(* IEC 61131-3 sources: plc-st-coding-agent/progress/evidence/f14_v11_public_20261113/jobs/codex_minimax-m27, 6 files *)

(* ---- public-easy-01.candidate_01.st ---- *)
(* ENGINEERING_CONTRACT
 * Filling Line State Machine - 6 states, sequential operation
 * PUB001: bottleSensor TRUE → Pump_Motor := TRUE (hold until cleaningConfirmButton)
 * PUB002: cleaningConfirmButton → Filling_Valve := TRUE (hold until fillingConfirmButton)
 * PUB003: fillingConfirmButton → Capping_Machine := TRUE (hold until cappingConfirmButton)
 * PUB004: cappingConfirmButton → Packing_Machine := TRUE (hold until packingConfirmButton)
 * PUB005: packingConfirmButton → Completion_Light := TRUE (hold until finishedButton)
 * PUB006: finishedButton → Completion_Light := FALSE; all outputs FALSE; reset to IDLE
 * State retention: outputs held until explicitly deactivated by state transition or reset
 * Reset priority: finishedButton (PUB006) clears all outputs and returns to IDLE
 *)

(* CONTRACT_RULES [] *)

FUNCTION_BLOCK FillingLineControl
VAR_INPUT
    bottleSensor          : BOOL;
    cleaningConfirmButton : BOOL;
    fillingConfirmButton  : BOOL;
    cappingConfirmButton  : BOOL;
    packingConfirmButton  : BOOL;
    finishedButton        : BOOL;
END_VAR
VAR_OUTPUT
    Pump_Motor      : BOOL;
    Filling_Valve   : BOOL;
    Capping_Machine : BOOL;
    Packing_Machine : BOOL;
    Completion_Light: BOOL;
END_VAR
VAR
    State : INT := 0;
END_VAR

// State machine: 0=IDLE, 1=CLEANING, 2=FILLING, 3=CAPPING, 4=PACKING, 5=COMPLETE
CASE State OF
    0: // IDLE - waiting for bottle
        Pump_Motor      := FALSE;
        Filling_Valve   := FALSE;
        Capping_Machine := FALSE;
        Packing_Machine := FALSE;
        Completion_Light:= FALSE;

        IF bottleSensor THEN
            State := 1;
        END_IF;

    1: // CLEANING
        Pump_Motor := TRUE;

        IF cleaningConfirmButton THEN
            Pump_Motor := FALSE;
            State := 2;
        END_IF;

    2: // FILLING
        Filling_Valve := TRUE;

        IF fillingConfirmButton THEN
            Filling_Valve := FALSE;
            State := 3;
        END_IF;

    3: // CAPPING
        Capping_Machine := TRUE;

        IF cappingConfirmButton THEN
            Capping_Machine := FALSE;
            State := 4;
        END_IF;

    4: // PACKING
        Packing_Machine := TRUE;

        IF packingConfirmButton THEN
            Packing_Machine := FALSE;
            State := 5;
        END_IF;

    5: // COMPLETE - bottle ready for pickup
        Completion_Light := TRUE;

        IF finishedButton THEN
            Completion_Light := FALSE;
            State := 0;
        END_IF;

END_CASE;

END_FUNCTION_BLOCK

(* ---- public-easy-01.raw_candidate_01.st ---- *)
(* ENGINEERING_CONTRACT
 * Filling Line State Machine - 6 states, sequential operation
 * PUB001: bottleSensor TRUE → Pump_Motor := TRUE (hold until cleaningConfirmButton)
 * PUB002: cleaningConfirmButton → Filling_Valve := TRUE (hold until fillingConfirmButton)
 * PUB003: fillingConfirmButton → Capping_Machine := TRUE (hold until cappingConfirmButton)
 * PUB004: cappingConfirmButton → Packing_Machine := TRUE (hold until packingConfirmButton)
 * PUB005: packingConfirmButton → Completion_Light := TRUE (hold until finishedButton)
 * PUB006: finishedButton → Completion_Light := FALSE; all outputs FALSE; reset to IDLE
 * State retention: outputs held until explicitly deactivated by state transition or reset
 * Reset priority: finishedButton (PUB006) clears all outputs and returns to IDLE
 *)

(* CONTRACT_RULES [] *)

FUNCTION_BLOCK FillingLineControl
VAR_INPUT
    bottleSensor          : BOOL;
    cleaningConfirmButton : BOOL;
    fillingConfirmButton  : BOOL;
    cappingConfirmButton  : BOOL;
    packingConfirmButton  : BOOL;
    finishedButton        : BOOL;
END_VAR
VAR_OUTPUT
    Pump_Motor      : BOOL;
    Filling_Valve   : BOOL;
    Capping_Machine : BOOL;
    Packing_Machine : BOOL;
    Completion_Light: BOOL;
END_VAR
VAR
    State : INT := 0;
END_VAR

// State machine: 0=IDLE, 1=CLEANING, 2=FILLING, 3=CAPPING, 4=PACKING, 5=COMPLETE
CASE State OF
    0: // IDLE - waiting for bottle
        Pump_Motor      := FALSE;
        Filling_Valve   := FALSE;
        Capping_Machine := FALSE;
        Packing_Machine := FALSE;
        Completion_Light:= FALSE;

        IF bottleSensor THEN
            State := 1;
        END_IF

    1: // CLEANING
        Pump_Motor := TRUE;

        IF cleaningConfirmButton THEN
            Pump_Motor := FALSE;
            State := 2;
        END_IF

    2: // FILLING
        Filling_Valve := TRUE;

        IF fillingConfirmButton THEN
            Filling_Valve := FALSE;
            State := 3;
        END_IF

    3: // CAPPING
        Capping_Machine := TRUE;

        IF cappingConfirmButton THEN
            Capping_Machine := FALSE;
            State := 4;
        END_IF

    4: // PACKING
        Packing_Machine := TRUE;

        IF packingConfirmButton THEN
            Packing_Machine := FALSE;
            State := 5;
        END_IF

    5: // COMPLETE - bottle ready for pickup
        Completion_Light := TRUE;

        IF finishedButton THEN
            Completion_Light := FALSE;
            State := 0;
        END_IF

END_CASE

END_FUNCTION_BLOCK

(* ---- public-easy-02.candidate_01.st ---- *)
(* ENGINEERING_CONTRACT
====================
PUB001: 76-318

State Retention:
- tmp_previous_value: RETAINED across scans (stores last cycle's DWORD value)
- All outputs: COMBINATIONAL (derived fresh each scan from current inputs + retained state)

Edge Detection Logic:
- Rising edge:  (current = 1) AND (previous = 0)  → risingBits = value & NOT previous
- Falling edge: (current = 0) AND (previous = 1)  → fallingBits = NOT value & previous
- Changed:      value <> previous

Counting:
- Count 1-bits in risingBits  → noOfRisingBits  (0-32)
- Count 1-bits in fallingBits → noOfFallingBits (0-32)

Priority:
- All outputs derived combinatorially in same scan
- No edge-only triggers or state machines

Units:
- risingBits/fallingBits: dimensionless bit patterns (DWORD)
- noOfRisingBits/noOfFallingBits: unsigned count (USINT, 0-32)
*)
FUNCTION_BLOCK FB_DualWordEdgeDetection
VAR
    tmp_previous_value : DWORD := 0;
END_VAR
VAR_OUTPUT
    hasChanged      : BOOL;
    hasRisingEdges  : BOOL;
    risingBits      : DWORD;
    noOfRisingBits  : USINT;
    hasFallingEdges : BOOL;
    fallingBits     : DWORD;
    noOfFallingBits : USINT;
END_VAR

risingBits  := value AND NOT tmp_previous_value;
fallingBits := NOT value AND tmp_previous_value;

hasChanged      := (value <> tmp_previous_value);
hasRisingEdges  := (risingBits <> 0);
hasFallingEdges := (fallingBits <> 0);

noOfRisingBits  := 0;
FOR i := 0 TO 31 DO
    IF SHR(risingBits, i) AND 1 = 1 THEN
        noOfRisingBits := noOfRisingBits + 1;
    END_IF;
END_FOR;

noOfFallingBits := 0;
FOR i := 0 TO 31 DO
    IF SHR(fallingBits, i) AND 1 = 1 THEN
        noOfFallingBits := noOfFallingBits + 1;
    END_IF;
END_FOR;

tmp_previous_value := value;
END_FUNCTION_BLOCK

(* ---- public-easy-02.candidate_02.st ---- *)
(* ENGINEERING_CONTRACT
====================
PUB001: 76-318

State Retention:
- tmp_previous_value: RETAINED across scans (stores last cycle's DWORD value)
- All outputs: COMBINATIONAL (derived fresh each scan from current inputs + retained state)

Edge Detection Logic:
- Rising edge:  (current = 1) AND (previous = 0)  → risingBits = value & NOT previous
- Falling edge: (current = 0) AND (previous = 1)  → fallingBits = NOT value & previous
- Changed:      value <> previous

Counting:
- Count 1-bits in risingBits  → noOfRisingBits  (0-32)
- Count 1-bits in fallingBits → noOfFallingBits (0-32)

Priority:
- All outputs derived combinatorially in same scan
- No edge-only triggers or state machines

Units:
- risingBits/fallingBits: dimensionless bit patterns (DWORD)
- noOfRisingBits/noOfFallingBits: unsigned count (USINT, 0-32)
*)
FUNCTION_BLOCK FB_DualWordEdgeDetection
VAR_INPUT
    value : DWORD;
END_VAR
VAR
    tmp_previous_value : DWORD := 0;
    i                  : INT;
    tmp_bit            : DWORD;
END_VAR
VAR_OUTPUT
    hasChanged      : BOOL;
    hasRisingEdges  : BOOL;
    risingBits      : DWORD;
    noOfRisingBits  : USINT;
    hasFallingEdges : BOOL;
    fallingBits     : DWORD;
    noOfFallingBits : USINT;
END_VAR

risingBits  := value AND NOT tmp_previous_value;
fallingBits := (NOT value) AND tmp_previous_value;

hasChanged      := (value <> tmp_previous_value);
hasRisingEdges  := (risingBits <> 0);
hasFallingEdges := (fallingBits <> 0);

noOfRisingBits := 0;
FOR i := 0 TO 31 DO
    tmp_bit := SHR(risingBits, i);
    IF TO_BOOL(tmp_bit AND 1) THEN
        noOfRisingBits := noOfRisingBits + 1;
    END_IF;
END_FOR;

noOfFallingBits := 0;
FOR i := 0 TO 31 DO
    tmp_bit := SHR(fallingBits, i);
    IF TO_BOOL(tmp_bit AND 1) THEN
        noOfFallingBits := noOfFallingBits + 1;
    END_IF;
END_FOR;

tmp_previous_value := value;
END_FUNCTION_BLOCK

(* ---- public-easy-02.raw_candidate_01.st ---- *)
(* ENGINEERING_CONTRACT
====================
PUB001: 76-318

State Retention:
- tmp_previous_value: RETAINED across scans (stores last cycle's DWORD value)
- All outputs: COMBINATIONAL (derived fresh each scan from current inputs + retained state)

Edge Detection Logic:
- Rising edge:  (current = 1) AND (previous = 0)  → risingBits = value & NOT previous
- Falling edge: (current = 0) AND (previous = 1)  → fallingBits = NOT value & previous
- Changed:      value <> previous

Counting:
- Count 1-bits in risingBits  → noOfRisingBits  (0-32)
- Count 1-bits in fallingBits → noOfFallingBits (0-32)

Priority:
- All outputs derived combinatorially in same scan
- No edge-only triggers or state machines

Units:
- risingBits/fallingBits: dimensionless bit patterns (DWORD)
- noOfRisingBits/noOfFallingBits: unsigned count (USINT, 0-32)
*)
FUNCTION_BLOCK FB_DualWordEdgeDetection
VAR
    tmp_previous_value : DWORD := 0;
END_VAR
VAR_OUTPUT
    hasChanged      : BOOL;
    hasRisingEdges  : BOOL;
    risingBits      : DWORD;
    noOfRisingBits  : USINT;
    hasFallingEdges : BOOL;
    fallingBits     : DWORD;
    noOfFallingBits : USINT;
END_VAR

risingBits  := value AND NOT tmp_previous_value;
fallingBits := NOT value AND tmp_previous_value;

hasChanged      := (value <> tmp_previous_value);
hasRisingEdges  := (risingBits <> 0);
hasFallingEdges := (fallingBits <> 0);

noOfRisingBits  := 0;
FOR i := 0 TO 31 DO
    IF SHR(risingBits, i) AND 1 = 1 THEN
        noOfRisingBits := noOfRisingBits + 1;
    END_IF;
END_FOR;

noOfFallingBits := 0;
FOR i := 0 TO 31 DO
    IF SHR(fallingBits, i) AND 1 = 1 THEN
        noOfFallingBits := noOfFallingBits + 1;
    END_IF;
END_FOR;

tmp_previous_value := value;
END_FUNCTION_BLOCK

(* ---- public-easy-02.raw_candidate_02.st ---- *)
(* ENGINEERING_CONTRACT
====================
PUB001: 76-318

State Retention:
- tmp_previous_value: RETAINED across scans (stores last cycle's DWORD value)
- All outputs: COMBINATIONAL (derived fresh each scan from current inputs + retained state)

Edge Detection Logic:
- Rising edge:  (current = 1) AND (previous = 0)  → risingBits = value & NOT previous
- Falling edge: (current = 0) AND (previous = 1)  → fallingBits = NOT value & previous
- Changed:      value <> previous

Counting:
- Count 1-bits in risingBits  → noOfRisingBits  (0-32)
- Count 1-bits in fallingBits → noOfFallingBits (0-32)

Priority:
- All outputs derived combinatorially in same scan
- No edge-only triggers or state machines

Units:
- risingBits/fallingBits: dimensionless bit patterns (DWORD)
- noOfRisingBits/noOfFallingBits: unsigned count (USINT, 0-32)
*)
FUNCTION_BLOCK FB_DualWordEdgeDetection
VAR_INPUT
    value : DWORD;
END_VAR
VAR
    tmp_previous_value : DWORD := 0;
    i                  : INT;
    tmp_bit            : DWORD;
END_VAR
VAR_OUTPUT
    hasChanged      : BOOL;
    hasRisingEdges  : BOOL;
    risingBits      : DWORD;
    noOfRisingBits  : USINT;
    hasFallingEdges : BOOL;
    fallingBits     : DWORD;
    noOfFallingBits : USINT;
END_VAR

risingBits  := value AND NOT tmp_previous_value;
fallingBits := (NOT value) AND tmp_previous_value;

hasChanged      := (value <> tmp_previous_value);
hasRisingEdges  := (risingBits <> 0);
hasFallingEdges := (fallingBits <> 0);

noOfRisingBits := 0;
FOR i := 0 TO 31 DO
    tmp_bit := SHR(risingBits, i);
    IF TO_BOOL(tmp_bit AND 1) THEN
        noOfRisingBits := noOfRisingBits + 1;
    END_IF;
END_FOR;

noOfFallingBits := 0;
FOR i := 0 TO 31 DO
    tmp_bit := SHR(fallingBits, i);
    IF TO_BOOL(tmp_bit AND 1) THEN
        noOfFallingBits := noOfFallingBits + 1;
    END_IF;
END_FOR;

tmp_previous_value := value;
END_FUNCTION_BLOCK
